Fanuc KAREL source: kt00599.KL

-- PROVISIONAL review KL for V770-1; original PC SHA256 afe23ec1703d367f3ed6ef422eb5a1a8f4eeea9d5dff7db565a37240e1735c6c
-- Incomplete behavior may be omitted. Consult companion uncertainty JSON. Do not deploy.
PROGRAM KT00599
%NOLOCKGROUP
VAR
  I1 : INTEGER
  I2 : INTEGER
  OUT : REAL
BEGIN
  -- UNRESOLVED_PC offsets 5-16; opcodes 2E,23
  -- UNRESOLVED_PC offsets 21-32; opcodes 2E,23
  -- UNRESOLVED_PC offsets 37-48; opcodes 2E,23
  -- UNRESOLVED_PC offsets 53-64; opcodes 2E,23
  -- UNRESOLVED_PC offsets 69-83; opcodes 21,48,64,23
  -- UNRESOLVED_PC offsets 88-92; opcodes 7F
END KT00599
